DATA_BLOCK "FRK_LineSource"
{ S7_Optimized_Access := 'TRUE' }
VERSION : 0.1
NON_RETAIN
VAR
    Image {ExternalAccessible := 'False'; ExternalVisible := 'False'; ExternalWritable := 'False'} : "ST_LineImage";
END_VAR
BEGIN
END_DATA_BLOCK
